Fanuc KAREL source: KT00003.KL

PROGRAM KT00003
%NOLOCKGROUP
VAR
  I1: INTEGER
  R2: REAL
  OUT: INTEGER
BEGIN
  I1 = 2
    R2 = 3.0
  OUT = I1 + R2
END KT00003
